// TIA Portal V18 export
FUNCTION "RESET_MODZONES" : Void   // FC10, LAD
{ S7_Optimized_Access := 'TRUE' }
// stored: SetENOAutomatically false
BEGIN

REGION Network 1: RESET MOD 1
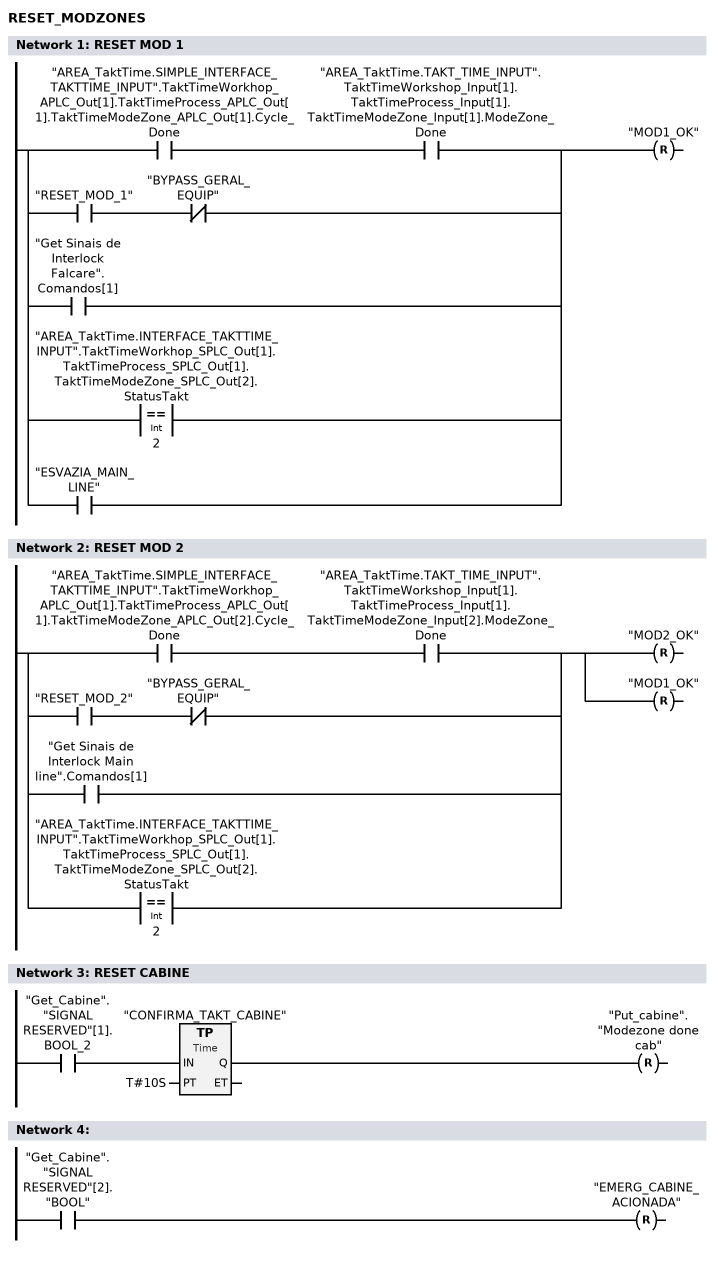
   RUNG wire#powerrail
      Contact( "AREA_TaktTime.SIMPLE_INTERFACE_TAKTTIME_INPUT".TaktTimeWorkhop_APLC_Out[1].TaktTimeProcess_APLC_Out[1].TaktTimeModeZone_APLC_Out[1].Cycle_Done )
      Contact( "AREA_TaktTime.TAKT_TIME_INPUT".TaktTimeWorkshop_Input[1].TaktTimeProcess_Input[1].TaktTimeModeZone_Input[1].ModeZone_Done )
      wire#w1
      R_Coil( "MOD1_OK" )
   END_RUNG
   RUNG wire#powerrail
      Contact( "RESET_MOD_1" )
      I_Contact( "BYPASS_GERAL_EQUIP" )
   END_RUNG wire#w1
   RUNG wire#powerrail
      Contact( "Get Sinais de Interlock Falcare".Comandos[1] )
   END_RUNG wire#w1
   RUNG wire#powerrail
      { S7_Templates := "SrcType := Int" } EQ_Contact(in1 := "AREA_TaktTime.INTERFACE_TAKTTIME_INPUT".TaktTimeWorkhop_SPLC_Out[1].TaktTimeProcess_SPLC_Out[1].TaktTimeModeZone_SPLC_Out[2].StatusTakt, in2 := 2)
   END_RUNG wire#w1
   RUNG wire#powerrail
      Contact( "ESVAZIA_MAIN_LINE" )
   END_RUNG wire#w1
   // the same network as SCL:
   IF ("AREA_TaktTime.SIMPLE_INTERFACE_TAKTTIME_INPUT".TaktTimeWorkhop_APLC_Out[1].TaktTimeProcess_APLC_Out[1].TaktTimeModeZone_APLC_Out[1].Cycle_Done AND "AREA_TaktTime.TAKT_TIME_INPUT".TaktTimeWorkshop_Input[1].TaktTimeProcess_Input[1].TaktTimeModeZone_Input[1].ModeZone_Done) OR ("RESET_MOD_1" AND NOT "BYPASS_GERAL_EQUIP") OR "Get Sinais de Interlock Falcare".Comandos[1] OR ("AREA_TaktTime.INTERFACE_TAKTTIME_INPUT".TaktTimeWorkhop_SPLC_Out[1].TaktTimeProcess_SPLC_Out[1].TaktTimeModeZone_SPLC_Out[2].StatusTakt = 2) OR "ESVAZIA_MAIN_LINE" THEN
       "MOD1_OK" := FALSE;
   END_IF;
END_REGION

REGION Network 2: RESET MOD 2
   RUNG wire#powerrail
      Contact( "AREA_TaktTime.SIMPLE_INTERFACE_TAKTTIME_INPUT".TaktTimeWorkhop_APLC_Out[1].TaktTimeProcess_APLC_Out[1].TaktTimeModeZone_APLC_Out[2].Cycle_Done )
      Contact( "AREA_TaktTime.TAKT_TIME_INPUT".TaktTimeWorkshop_Input[1].TaktTimeProcess_Input[1].TaktTimeModeZone_Input[2].ModeZone_Done )
      wire#w1
      R_Coil( "MOD2_OK" )
   END_RUNG
   RUNG wire#powerrail
      Contact( "RESET_MOD_2" )
      I_Contact( "BYPASS_GERAL_EQUIP" )
   END_RUNG wire#w1
   RUNG wire#powerrail
      Contact( "Get Sinais de Interlock Main line".Comandos[1] )
   END_RUNG wire#w1
   RUNG wire#powerrail
      { S7_Templates := "SrcType := Int" } EQ_Contact(in1 := "AREA_TaktTime.INTERFACE_TAKTTIME_INPUT".TaktTimeWorkhop_SPLC_Out[1].TaktTimeProcess_SPLC_Out[1].TaktTimeModeZone_SPLC_Out[2].StatusTakt, in2 := 2)
   END_RUNG wire#w1
   RUNG wire#w1
      R_Coil( "MOD1_OK" )
   END_RUNG
   // the same network as SCL:
   IF ("AREA_TaktTime.SIMPLE_INTERFACE_TAKTTIME_INPUT".TaktTimeWorkhop_APLC_Out[1].TaktTimeProcess_APLC_Out[1].TaktTimeModeZone_APLC_Out[2].Cycle_Done AND "AREA_TaktTime.TAKT_TIME_INPUT".TaktTimeWorkshop_Input[1].TaktTimeProcess_Input[1].TaktTimeModeZone_Input[2].ModeZone_Done) OR ("RESET_MOD_2" AND NOT "BYPASS_GERAL_EQUIP") OR "Get Sinais de Interlock Main line".Comandos[1] OR ("AREA_TaktTime.INTERFACE_TAKTTIME_INPUT".TaktTimeWorkhop_SPLC_Out[1].TaktTimeProcess_SPLC_Out[1].TaktTimeModeZone_SPLC_Out[2].StatusTakt = 2) THEN
       "MOD2_OK" := FALSE;
       "MOD1_OK" := FALSE;
   END_IF;
END_REGION

REGION Network 3: RESET CABINE
   RUNG wire#powerrail
      Contact( "Get_Cabine"."SIGNAL RESERVED"[1].BOOL_2 )
      { S7_Templates := "time_type := Time" } "CONFIRMA_TAKT_CABINE".TP(pt := T#10S, et =>)
      R_Coil( "Put_cabine"."Modezone done cab" )
   END_RUNG
   // the same network as SCL:
   "CONFIRMA_TAKT_CABINE".TP(IN := "Get_Cabine"."SIGNAL RESERVED"[1].BOOL_2, PT := T#10S);
   IF "CONFIRMA_TAKT_CABINE".Q THEN "Put_cabine"."Modezone done cab" := FALSE; END_IF;
END_REGION

REGION Network 4
   RUNG wire#powerrail
      Contact( "Get_Cabine"."SIGNAL RESERVED"[2]."BOOL" )
      R_Coil( "EMERG_CABINE_ACIONADA" )
   END_RUNG
   // the same network as SCL:
   IF "Get_Cabine"."SIGNAL RESERVED"[2]."BOOL" THEN "EMERG_CABINE_ACIONADA" := FALSE; END_IF;
END_REGION
END_FUNCTION
